TYPE ST_PolarIIChamber_CupLiftServiceStatus :
STRUCT
	JogPositive : ST_ServiceStatus;
	JogNegative : ST_ServiceStatus;
	IncrementalJog : ST_ServiceStatus;
	DecoupleStop : ST_ServiceStatus; // NaturalCompletion.
	TopPos : ST_ServiceStatus;
	MiddlePos : ST_ServiceStatus;
	DownPos : ST_ServiceStatus;
END_STRUCT
END_TYPE

(* stored: Version 1.1.0.1, ProductVersion 3.1.4026.18
   DUT ST_PolarIIChamber_CupLiftServiceStatus: Id {14000000-0000-0000-0000-000000000039} *)
